// TIA Portal V17 export
FUNCTION_BLOCK "FB_T04b_TON_Multi"   // FB142, LAD
{ S7_Optimized_Access := 'TRUE' }
// stored: IsIECCheckEnabled false, MemoryReserve 100, SetENOAutomatically false
   VAR_INPUT
      Demarrer : Bool;
      Duree : Time;
   END_VAR
   VAR_OUTPUT
      Tempo_OK : Bool;
      Ecoule : Time;
   END_VAR
   VAR
      tonDelai : TON_TIME;
   END_VAR
BEGIN

REGION Network 1: TON multi-instance
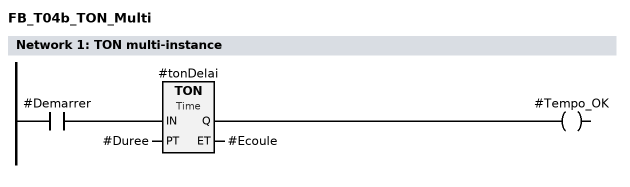
   RUNG wire#powerrail
      Contact( #Demarrer )
      { S7_Templates := "time_type := Time" } #tonDelai.TON(pt := #Duree, et => #Ecoule)
      Coil( #Tempo_OK )
   END_RUNG
   // the same network as SCL:
   #tonDelai(IN := #Demarrer, PT := #Duree, ET => #Ecoule);   // TON
   #Tempo_OK := #tonDelai.Q;
END_REGION
END_FUNCTION_BLOCK
